(*~
	<docu>
		<summary>
			KUKA robot controller running KSS / iiQKA.OS2 9.3 (ECat).
			The interface uses 64 input and 64 output bytes. Compared to TcoKrc4 v5 it adds LocalEstopOk, NormalStop,
			CutEnableDrives, user data in both directions and a new start sequence (interface is activated first,
			drives are switched on only when CutEnableDrives is present).
		</summary>
	</docu>
~*)
FUNCTION_BLOCK TcoKukaKssEcat_v_9_3_x EXTENDS TcoIo.TcoEcatComponent IMPLEMENTS TcoAbstractions.ITcoRobotics
VAR_INPUT
    inEnable : BOOL;
END_VAR
VAR_OUTPUT
END_VAR
VAR_IN_OUT
    inoData : TcoKukaKssEcat_IO_v_9_3_x;
END_VAR
VAR
	{attribute addProperty Name "<#Status#>"}
    {attribute clr [ReadOnly()]}
    _status : TcoKukaKss_Status_v_9_3_x;
	{attribute addProperty Name "<#Control#>"}
	_control : TcoKukaKss_Control_v_9_3_x;
	{attribute addProperty Name "<#Config#>"}
    _config : TcoKukaKss_Config_v_9_3_x;
	{attribute addProperty Name "<#ECat Error#>"}
    {attribute clr [ReadOnly()]}
    _busError : BOOL;

	_someTaskIsActive : BOOL;
	_stopTasksAreActive : BOOL;

	_reportTimer : TON;
	_errorReportTimer : TON;
	{attribute 'hide'}
	_manualPV : BOOL;
END_VAR
VAR
	{attribute addProperty Name "<#Start at Main#>"}
	_startAtMainTask : TcoKukaKss_StartAtMainTask_v_9_3_x(THIS^);

	{attribute addProperty Name "<#Start motors and program#>"}
	_startMotorsAndProgramTask : TcoKukaKss_StartMotorsAndProgramTask_v_9_3_x(THIS^);

	{attribute addProperty Name "<#Start program#>"}
	_startProgramTask : TcoKukaKss_StartProgramTask_v_9_3_x(THIS^);

	{attribute addProperty Name "<#Start motors#>"}
	_startMotorsTask : TcoKukaKss_StartMotorsTask_v_9_3_x(THIS^);

	{attribute addProperty Name "<#Start movements#>"}
	_startMovementsTask : TcoKukaKss_StartMovementsTask_v_9_3_x(THIS^);

	{attribute addProperty Name "<#Start motors program and movements#>"}
	_startMotorsProgramAndMovementsTask : TcoKukaKss_StartMotorsProgramAndMovementsTask_v_9_3_x(THIS^);

	{attribute addProperty Name "<#Stop movements#>"}
	_stopMovementsTask : TcoKukaKss_StopMovementsTask_v_9_3_x(THIS^);

	{attribute addProperty Name "<#Stop movenents and program#>"}
	_stopMovementsAndProgramTask : TcoKukaKss_StopMovementsAndProgramTask_v_9_3_x(THIS^);

	{attribute addProperty Name "<#Stop program#>"}
	_stopProgramTask : TcoKukaKss_StopProgramTask_v_9_3_x(THIS^);

	{attribute addProperty Name "<#Stop motors#>"}
	_stopMotorsTask : TcoKukaKss_StopMotorsTask_v_9_3_x(THIS^);

	{attribute addProperty Name "<#Reset all outputs#>"}
	_resetAllOutputsTask : TcoKukaKss_ResetAllOutputsTask_v_9_3_x(THIS^);

    {attribute addProperty Name "<#Restore#>"}
    _restoreTask : TcoCore.TcoTask(THIS^);
END_VAR

IF NOT __ISVALIDREF(inoData) THEN
    Messenger.Post('Invalid reference', TcoCore.eMessageCategory.ProgrammingError);
    RETURN;
END_IF

SUPER^(AdsAddr := AdsAddr);
_busError := NOT SUPER^._ecatState.EcatOk;

UpdateStatus();

//MoveEnable follows the manual mode: set on entering manual mode, reset on leaving it
IF _status.State.Manual AND NOT _manualPV THEN
    _control.MoveEnable := TRUE;
ELSIF NOT _status.State.Manual AND _manualPV THEN
    _control.MoveEnable := FALSE;
END_IF
_manualPV := _status.State.Manual;

_stopTasksAreActive := _stopMovementsTask.Busy OR _stopMovementsAndProgramTask.Busy OR _stopProgramTask.Busy OR _stopMotorsTask.Busy;

_startAtMainTask.Enabled := NOT _stopTasksAreActive;
_startAtMainTask(inoConfig := _config, inoControl := _control, inoStatus := _status);

_startProgramTask.Enabled := NOT _stopTasksAreActive AND NOT _startMotorsAndProgramTask.Busy AND NOT _startMotorsTask.Busy;
_startProgramTask(inoConfig := _config, inoControl := _control, inoStatus := _status);

_startMotorsTask.Enabled := NOT _stopTasksAreActive AND NOT _startMotorsProgramAndMovementsTask.Busy AND NOT _startMotorsAndProgramTask.Busy AND NOT _startProgramTask.Busy;
_startMotorsTask(inoConfig := _config, inoControl := _control, inoStatus := _status);

_startMotorsAndProgramTask.Enabled := NOT _stopTasksAreActive AND NOT _startProgramTask.Busy AND NOT _startMotorsTask.Busy;
_startMotorsAndProgramTask(inoConfig := _config, inoControl := _control, inoStatus := _status);

_startMovementsTask.Enabled := NOT _startMotorsProgramAndMovementsTask.Busy AND NOT _stopMotorsTask.Busy;
_startMovementsTask(inoConfig := _config, inoControl := _control, inoStatus := _status);

_startMotorsProgramAndMovementsTask.Enabled := NOT _startMovementsTask.Busy AND NOT _stopMotorsTask.Busy;
_startMotorsProgramAndMovementsTask(refStartMotorsAndProgramTask := _startMotorsAndProgramTask,
    inoConfig := _config,
    inoControl := _control,
    inoStatus := _status);

_stopMovementsTask.Enabled := TRUE;
_stopMovementsTask(inoConfig := _config, inoControl := _control, inoStatus := _status);

_stopMotorsTask.Enabled := TRUE;
_stopMotorsTask(inoConfig := _config, inoControl := _control, inoStatus := _status);

_stopProgramTask.Enabled := TRUE;
_stopProgramTask(inoConfig := _config, inoControl := _control, inoStatus := _status);

_stopMovementsAndProgramTask.Enabled := TRUE;
_stopMovementsAndProgramTask(inoConfig := _config, inoControl := _control, inoStatus := _status);

_someTaskIsActive := _startAtMainTask.Busy OR
    _startProgramTask.Busy OR
    _startMotorsTask.Busy OR
    _startMotorsAndProgramTask.Busy OR
    _startMovementsTask.Busy OR
    _startMotorsProgramAndMovementsTask.Busy OR
    _stopMovementsTask.Busy OR
    _stopMovementsAndProgramTask.Busy OR
    _stopProgramTask.Busy OR
    _stopMotorsTask.Busy;

_resetAllOutputsTask.Enabled := NOT _someTaskIsActive;
_resetAllOutputsTask(inoConfig := _config, inoControl := _control, inoStatus := _status);

//*************RESTORE********************
_restoreTask.Enabled := TRUE;
IF _restoreTask.Execute() THEN
    Restore();
    _restoreTask.DoneWhen(TRUE);
END_IF
//****************************************

//do not publish diagnostic message when component is not used
IF _someTaskIsActive THEN
    IF NOT _status.State.AlarmStopActive THEN
        Messenger.Error('<#Emergency stop active#>');
    END_IF;
    IF NOT _status.State.LocalEstopOk THEN
        Messenger.Error('<#Local emergency stop active#>');
    END_IF;
    IF NOT _status.State.UserSafetySwitchClosed THEN
        Messenger.Warning('<#Safety Error #>');
    END_IF;
END_IF;

_errorReportTimer(IN := _status.State.Error, PT := _config.InfoTime);
Messenger.OnCondition(_errorReportTimer.Q).Error(_sb.Clear()
        .Append('<#Robot reported an error: #>')
        .Append(UDINT_TO_STRING(_status.State.EventId))
        .Append(' |[[0]AdvancedDiagnosticMessage]|')
        .Append('.')
        .Append('For details see the service mode')
        .ToString());

_reportTimer(IN := _status.State.Manual, PT := _config.InfoTime);
Messenger.OnCondition(_reportTimer.Q).Warning('<#Robot in manual mode. MoveEnable is set on entering manual mode!#>');

UpdateControl();

(*~
	<docu>
		<summary>
			Gets the configuration of the robot. 					
		</summary>			
	</docu>	
~*)
PROPERTY Config : REFERENCE TO TcoKukaKss_Config_v_9_3_x
GET
Config REF= _config;
END_GET
END_PROPERTY

PROPERTY PUBLIC Control : REFERENCE TO TcoKukaKss_Control_v_9_3_x
GET
Control REF= _control;
END_GET
END_PROPERTY

(*~
	<docu>
		<summary>
			Gets the status of the robot. 					
		</summary>			
	</docu>	
~*)
PROPERTY Status : REFERENCE TO TcoKukaKss_Status_v_9_3_x
GET
Status REF= _status;
END_GET
END_PROPERTY

METHOD FB_init : BOOL
VAR_INPUT
	bInitRetains : BOOL; // if TRUE, the retain variables are initialized (warm start / cold start)
	bInCopyCode : BOOL;  // if TRUE, the instance afterwards gets moved into the copy code (online change)
  	ParentObject : ITcoObject;	
END_VAR
END_METHOD

(*~
	<docu>
		<summary>
			Restores this instance to the Ready state. Can be called explicitly or from within one of the restore mechanisms.	
		</summary>			
	</docu>	
~*)
METHOD Restore : ITcoRestorable
RestoreTasks();

_control.GlobalSpeed := 0;
_control.ActivateInterface := FALSE;
_control.ErrorConfirmation := FALSE;
_control.ExternalStart := FALSE;
_control.MasterMode := 0;
_control.ToolNo := 0;
_control.WorkobjectNo := 0;
_control.PointNo := 0;
_control.UserSpecSpeed1 := 0;
_control.UserSpecSpeed2 := 0;
_control.Coordinates.X := 0;
_control.Coordinates.Y := 0;
_control.Coordinates.Z := 0;
_control.Coordinates.Rx := 0;
_control.Coordinates.Ry := 0;
_control.Coordinates.Rz := 0;
END_METHOD

METHOD INTERNAL RestoreTasks
_startAtMainTask.Restore();
_startMotorsAndProgramTask.Restore();
_startProgramTask.Restore();
_startMotorsTask.Restore();
_startMovementsTask.Restore();
_startMotorsProgramAndMovementsTask.Restore();
_stopMovementsTask.Restore();
_stopMovementsAndProgramTask.Restore();
_stopProgramTask.Restore();
_stopMotorsTask.Restore();
_resetAllOutputsTask.Restore();
END_METHOD

(*~
	<docu>
		<summary>
		    Custom service (manual, maintenance) logic.
			This method must be implemented in derived class.
		</summary>			
	</docu>	
~*)
METHOD PROTECTED ServiceMode
END_METHOD

METHOD PUBLIC StartAtMain : TcoCore.ITcoTaskStatus
StartAtMain := _startAtMainTask.Invoke();
END_METHOD

PROPERTY StartAtMainTask : TcoCore.ITcoTaskStatus
GET
StartAtMainTask := _startAtMainTask;
END_GET
END_PROPERTY

METHOD PUBLIC StartMotors : TcoCore.ITcoTaskStatus
StartMotors := _startMotorsTask.Invoke();
END_METHOD

PROPERTY StartMotorsTask : TcoCore.ITcoTaskStatus
GET
StartMotorsTask := _startMotorsTask;
END_GET
END_PROPERTY

METHOD PUBLIC StartMotorsAndProgram : TcoCore.ITcoTaskStatus
StartMotorsAndProgram := _startMotorsAndProgramTask.Invoke();
END_METHOD

PROPERTY StartMotorsAndProgramTask : TcoCore.ITcoTaskStatus
GET
StartMotorsAndProgramTask := _startMotorsAndProgramTask;
END_GET
END_PROPERTY

METHOD PUBLIC StartProgram : TcoCore.ITcoTaskStatus
StartProgram := _startProgramTask.Invoke();
END_METHOD

PROPERTY StartProgramTask : TcoCore.ITcoTaskStatus
GET
StartProgramTask := _startProgramTask;
END_GET
END_PROPERTY

METHOD PUBLIC StartMovements : TcoCore.ITcoTaskStatus
VAR_INPUT
	inData : TcoRoboticsMovementsParams;
END_VAR
StartMovements := _startMovementsTask.InvokeWithParams(inData);
END_METHOD

PROPERTY StartMovementsTask : TcoCore.ITcoTaskStatus
GET
StartMovementsTask := _startMovementsTask;
END_GET
END_PROPERTY

METHOD PUBLIC StartMotorsProgramAndMovements : TcoCore.ITcoTaskStatus
VAR_INPUT
	inData : TcoRoboticsMovementsParams;
END_VAR
StartMotorsProgramAndMovements := _startMotorsProgramAndMovementsTask.InvokeWithParams(inData);
END_METHOD

PROPERTY StartMotorsProgramAndMovementsTask : TcoCore.ITcoTaskStatus
GET
StartMotorsProgramAndMovementsTask := _startMotorsProgramAndMovementsTask;
END_GET
END_PROPERTY

METHOD PUBLIC StopMotors : TcoCore.ITcoTaskStatus
StopMotors := _stopMotorsTask.Invoke();
END_METHOD

PROPERTY StopMotorsTask : TcoCore.ITcoTaskStatus
GET
StopMotorsTask := _stopMotorsTask;
END_GET
END_PROPERTY

METHOD PUBLIC StopMovements : TcoCore.ITcoTaskStatus
VAR_INPUT
	inStopType : eTcoRoboticsStopType;
END_VAR
StopMovements := _stopMovementsTask.InvokeWithParams(inStopType);
END_METHOD

PROPERTY StopMovementsTask : TcoCore.ITcoTaskStatus
GET
StopMovementsTask := _stopMovementsTask;
END_GET
END_PROPERTY

METHOD PUBLIC StopMovementsAndProgram : TcoCore.ITcoTaskStatus
VAR_INPUT
	inStopType : eTcoRoboticsStopType;
END_VAR
StopMovementsAndProgram := _stopMovementsAndProgramTask.InvokeWithParams(inStopType);
END_METHOD

PROPERTY StopMovementsAndProgramTask : TcoCore.ITcoTaskStatus
GET
StopMovementsAndProgramTask := _stopMovementsAndProgramTask;
END_GET
END_PROPERTY

METHOD PUBLIC StopProgram : TcoCore.ITcoTaskStatus
StopProgram := _stopProgramTask.Invoke();
END_METHOD

PROPERTY StopProgramTask : TcoCore.ITcoTaskStatus
GET
StopProgramTask := _stopProgramTask;
END_GET
END_PROPERTY

METHOD PUBLIC ResetAllOutputs : TcoCore.ITcoTaskStatus
ResetAllOutputs := _resetAllOutputsTask.Invoke();
END_METHOD

PROPERTY ResetAllOutputsTask : TcoCore.ITcoTaskStatus
GET
ResetAllOutputsTask := _resetAllOutputsTask;
END_GET
END_PROPERTY

METHOD INTERNAL UpdateControl
VAR
	index : INT;
END_VAR
//SYSTEM OUTPUTS
index:=0;
inoData.Out.Outputs[index].0 := _control.ExternalStart;
inoData.Out.Outputs[index].1 := _control.MoveEnable;
inoData.Out.Outputs[index].2 := _control.ErrorConfirmation;
inoData.Out.Outputs[index].3 := _control.DrivesOff;
inoData.Out.Outputs[index].4 := _control.DrivesOn;
inoData.Out.Outputs[index].5 := _control.ActivateInterface;
inoData.Out.Outputs[index].6 := _control.StartAtMain;
inoData.Out.Outputs[index].7 := FALSE;
index:=1;
inoData.Out.Outputs[index] := 0;

//Tool signals
index:=2;
inoData.Out.Outputs[index].0 := _control.Tool_1_Retract;
inoData.Out.Outputs[index].1 := _control.Tool_1_Extend;
inoData.Out.Outputs[index].2 := _control.Tool_2_Retract;
inoData.Out.Outputs[index].3 := _control.Tool_2_Extend;
inoData.Out.Outputs[index].4 := _control.Tool_3_Retract;
inoData.Out.Outputs[index].5 := _control.Tool_3_Extend;
inoData.Out.Outputs[index].6 := _control.Tool_4_Retract;
inoData.Out.Outputs[index].7 := _control.Tool_4_Extend;
//master mode such as manual/auto ....
index:=3;
inoData.Out.Outputs[index] := _control.MasterMode;
//zone
index:=5;
inoData.Out.Outputs[index] := _control.Zone;
//position
index:=6;
inoData.Out.Outputs[index] := _control.InPosition;

//Movement parameters
index:=7;
inoData.Out.Outputs[index] := _control.ActionNo;
index:=8;
inoData.Out.Outputs[index] := _control.GlobalSpeed;
index:=9;
inoData.Out.Outputs[index] := _control.ToolNo;
index:=10;
inoData.Out.Outputs[index] := _control.WorkobjectNo;
index:=11;
inoData.Out.Outputs[index] := _control.PointNo;
index:=12;
TcoUtilities.TcoDintToBytes(inFormat:=TcoUtilities.eTcoDataFormat.LittleEndian,
							inValue:=REAL_TO_DINT(_control.UserSpecSpeed1),
							outByte0:=inoData.Out.Outputs[index],
							outByte1:=inoData.Out.Outputs[index+1],
							outByte2:=inoData.Out.Outputs[index+2],
							outByte3:=inoData.Out.Outputs[index+3]);
index:=16;
TcoUtilities.TcoDintToBytes(inFormat:=TcoUtilities.eTcoDataFormat.LittleEndian,
							inValue:=REAL_TO_DINT(_control.UserSpecSpeed2),
							outByte0:=inoData.Out.Outputs[index],
							outByte1:=inoData.Out.Outputs[index+1],
							outByte2:=inoData.Out.Outputs[index+2],
							outByte3:=inoData.Out.Outputs[index+3]);

//Coordinates
index:=20;
TcoUtilities.TcoDintToBytes(inFormat:=TcoUtilities.eTcoDataFormat.LittleEndian,
							inValue:=REAL_TO_DINT(_control.Coordinates.X * 10000.0),
							outByte0:=inoData.Out.Outputs[index],
							outByte1:=inoData.Out.Outputs[index+1],
							outByte2:=inoData.Out.Outputs[index+2],
							outByte3:=inoData.Out.Outputs[index+3]);
index:=24;
TcoUtilities.TcoDintToBytes(inFormat:=TcoUtilities.eTcoDataFormat.LittleEndian,
							inValue:=REAL_TO_DINT(_control.Coordinates.Y * 10000.0),
							outByte0:=inoData.Out.Outputs[index],
							outByte1:=inoData.Out.Outputs[index+1],
							outByte2:=inoData.Out.Outputs[index+2],
							outByte3:=inoData.Out.Outputs[index+3]);
index:=28;
TcoUtilities.TcoDintToBytes(inFormat:=TcoUtilities.eTcoDataFormat.LittleEndian,
							inValue:=REAL_TO_DINT(_control.Coordinates.Z * 10000.0),
							outByte0:=inoData.Out.Outputs[index],
							outByte1:=inoData.Out.Outputs[index+1],
							outByte2:=inoData.Out.Outputs[index+2],
							outByte3:=inoData.Out.Outputs[index+3]);
index:=32;
TcoUtilities.TcoDintToBytes(inFormat:=TcoUtilities.eTcoDataFormat.LittleEndian,
							inValue:=REAL_TO_DINT(_control.Coordinates.Rx * 10000.0),
							outByte0:=inoData.Out.Outputs[index],
							outByte1:=inoData.Out.Outputs[index+1],
							outByte2:=inoData.Out.Outputs[index+2],
							outByte3:=inoData.Out.Outputs[index+3]);
index:=36;
TcoUtilities.TcoDintToBytes(inFormat:=TcoUtilities.eTcoDataFormat.LittleEndian,
							inValue:=REAL_TO_DINT(_control.Coordinates.Ry * 10000.0),
							outByte0:=inoData.Out.Outputs[index],
							outByte1:=inoData.Out.Outputs[index+1],
							outByte2:=inoData.Out.Outputs[index+2],
							outByte3:=inoData.Out.Outputs[index+3]);
index:=40;
TcoUtilities.TcoDintToBytes(inFormat:=TcoUtilities.eTcoDataFormat.LittleEndian,
							inValue:=REAL_TO_DINT(_control.Coordinates.Rz * 10000.0),
							outByte0:=inoData.Out.Outputs[index],
							outByte1:=inoData.Out.Outputs[index+1],
							outByte2:=inoData.Out.Outputs[index+2],
							outByte3:=inoData.Out.Outputs[index+3]);

//User data from PLC to robot
FOR index := 0 TO 19 DO
	inoData.Out.Outputs[44 + index] := _control.DataToRobot[index];
END_FOR
END_METHOD

METHOD INTERNAL UpdateStatus
VAR
	index : INT;
	_bytes : DINT;
END_VAR
//SYSTEM INPUTS
index:=0;
_status.State.RcReady := inoData.In.Inputs[index].0;
_status.State.AlarmStopActive := inoData.In.Inputs[index].1;
_status.State.UserSafetySwitchClosed := inoData.In.Inputs[index].2;
_status.State.DrivesReady := inoData.In.Inputs[index].3;
_status.State.RobotCalibrated := inoData.In.Inputs[index].4;
_status.State.InterfaceActivated := inoData.In.Inputs[index].5;
_status.State.StopMess := inoData.In.Inputs[index].6;
_status.State.RobotStopped := inoData.In.Inputs[index].7;

index:=1;
_status.State.InHome := inoData.In.Inputs[index].0;
_status.State.Manual := inoData.In.Inputs[index].1;
_status.State.LocalEstopOk := inoData.In.Inputs[index].2;
_status.State.ExternalAutomatic := inoData.In.Inputs[index].3;
_status.State.ProActive := inoData.In.Inputs[index].4;
_status.State.PpMoved := inoData.In.Inputs[index].5;
_status.State.Error := inoData.In.Inputs[index].6;
_status.State.ProgramMoveActive := inoData.In.Inputs[index].7;

//Area/positions flags this should be obsolete because Zones and InPosition is used as byte below
index:=2;
_status.State.InArea_1 := inoData.In.Inputs[index].0;
_status.State.InArea_2 := inoData.In.Inputs[index].1;
_status.State.InArea_3 := inoData.In.Inputs[index].2;
_status.State.InArea_4 := inoData.In.Inputs[index].3;
_status.State.InPosition_1 := inoData.In.Inputs[index].4;
_status.State.InPosition_2 := inoData.In.Inputs[index].5;
_status.State.InPosition_3 := inoData.In.Inputs[index].6;
_status.State.InPosition_4 := inoData.In.Inputs[index].7;

//Tool signals
index:=3;
_status.State.Tool_1_Retract := inoData.In.Inputs[index].0;
_status.State.Tool_1_Extend := inoData.In.Inputs[index].1;
_status.State.Tool_2_Retract := inoData.In.Inputs[index].2;
_status.State.Tool_2_Extend := inoData.In.Inputs[index].3;
_status.State.Tool_3_Retract := inoData.In.Inputs[index].4;
_status.State.Tool_3_Extend := inoData.In.Inputs[index].5;
_status.State.Tool_4_Retract := inoData.In.Inputs[index].6;
_status.State.Tool_4_Extend := inoData.In.Inputs[index].7;

//Normal stop / drives enable (KSS 9.3)
index:=4;
_status.State.NormalStop := inoData.In.Inputs[index].0;
_status.State.CutEnableDrives := inoData.In.Inputs[index].1;

index:=5;
_status.State.Zone := inoData.In.Inputs[index];
index:=6;
_status.State.InPosition := inoData.In.Inputs[index];

//Movement parameters
index:=7;
_status.State.ActionNo := inoData.In.Inputs[index];
index:=8;
_status.State.GlobalSpeed := inoData.In.Inputs[index];
index:=9;
_status.State.ToolNo := inoData.In.Inputs[index];
index:=10;
_status.State.WorkobjectNo := inoData.In.Inputs[index];
index:=11;
_status.State.PointNo := inoData.In.Inputs[index];
index:=12;
_status.State.UserSpecSpeed1 := TcoUtilities.TcoBytesToDint(inFormat:=TcoUtilities.eTcoDataFormat.LittleEndian,
							inByte0:=inoData.In.Inputs[index],
							inByte1:=inoData.In.Inputs[index+1],
							inByte2:=inoData.In.Inputs[index+2],
							inByte3:=inoData.In.Inputs[index+3]);
index:=16;
_status.State.UserSpecSpeed2 := TcoUtilities.TcoBytesToDint(inFormat:=TcoUtilities.eTcoDataFormat.LittleEndian,
							inByte0:=inoData.In.Inputs[index],
							inByte1:=inoData.In.Inputs[index+1],
							inByte2:=inoData.In.Inputs[index+2],
							inByte3:=inoData.In.Inputs[index+3]);
index:=20;
_bytes := TcoUtilities.TcoBytesToDint(inFormat:=TcoUtilities.eTcoDataFormat.LittleEndian,
							inByte0:=inoData.In.Inputs[index],
							inByte1:=inoData.In.Inputs[index+1],
							inByte2:=inoData.In.Inputs[index+2],
							inByte3:=inoData.In.Inputs[index+3]);
_status.State.Coordinates.X := DINT_TO_REAL(_bytes) / 10000.0;

index:=24;
_bytes := TcoUtilities.TcoBytesToDint(inFormat:=TcoUtilities.eTcoDataFormat.LittleEndian,
							inByte0:=inoData.In.Inputs[index],
							inByte1:=inoData.In.Inputs[index+1],
							inByte2:=inoData.In.Inputs[index+2],
							inByte3:=inoData.In.Inputs[index+3]);
_status.State.Coordinates.Y := DINT_TO_REAL(_bytes) / 10000.0;

index:=28;
_bytes := TcoUtilities.TcoBytesToDint(inFormat:=TcoUtilities.eTcoDataFormat.LittleEndian,
							inByte0:=inoData.In.Inputs[index],
							inByte1:=inoData.In.Inputs[index+1],
							inByte2:=inoData.In.Inputs[index+2],
							inByte3:=inoData.In.Inputs[index+3]);
_status.State.Coordinates.Z := DINT_TO_REAL(_bytes) / 10000.0;

index:=32;
_bytes := TcoUtilities.TcoBytesToDint(inFormat:=TcoUtilities.eTcoDataFormat.LittleEndian,
							inByte0:=inoData.In.Inputs[index],
							inByte1:=inoData.In.Inputs[index+1],
							inByte2:=inoData.In.Inputs[index+2],
							inByte3:=inoData.In.Inputs[index+3]);
_status.State.Coordinates.Rx := DINT_TO_REAL(_bytes) / 10000.0;

index:=36;
_bytes := TcoUtilities.TcoBytesToDint(inFormat:=TcoUtilities.eTcoDataFormat.LittleEndian,
							inByte0:=inoData.In.Inputs[index],
							inByte1:=inoData.In.Inputs[index+1],
							inByte2:=inoData.In.Inputs[index+2],
							inByte3:=inoData.In.Inputs[index+3]);
_status.State.Coordinates.Ry := DINT_TO_REAL(_bytes) / 10000.0;

index:=40;
_bytes := TcoUtilities.TcoBytesToDint(inFormat:=TcoUtilities.eTcoDataFormat.LittleEndian,
							inByte0:=inoData.In.Inputs[index],
							inByte1:=inoData.In.Inputs[index+1],
							inByte2:=inoData.In.Inputs[index+2],
							inByte3:=inoData.In.Inputs[index+3]);
_status.State.Coordinates.Rz := DINT_TO_REAL(_bytes) / 10000.0;

index:=44;
_status.State.EventId := TcoUtilities.TcoBytesToUDint(inFormat:=TcoUtilities.eTcoDataFormat.LittleEndian,
							inByte0:=inoData.In.Inputs[index],
							inByte1:=inoData.In.Inputs[index+1],
							inByte2:=inoData.In.Inputs[index+2],
							inByte3:=inoData.In.Inputs[index+3]);

//User data from robot to PLC
FOR index := 0 TO 15 DO
	_status.State.DataFromRobot[index] := inoData.In.Inputs[48 + index];
END_FOR
END_METHOD

END_FUNCTION_BLOCK

(* stored: Version 1.1.0.1, ProductVersion 3.1.4024.12
   POU TcoKukaKssEcat_v_9_3_x: Id {8240f261-28f6-44a7-bcaa-32d5ed3116a8}, SpecialFunc None
   Folder Operations: Id {027f61ae-e71f-4a4c-8c22-228286bc5d5f}
   Folder Task: Id {2c37f829-6297-4777-bc3f-0fc886118850}
   Property Config: Id {4d37f924-eb41-4fef-9edc-76d0b4f40692}
   Get Get: Id {2258dc20-4fdb-45fe-b63a-6505710d1a93}
   Property Control: Id {e3180703-86e2-43b3-b541-81614d7caa3a}
   Get Get: Id {5ec5fc1e-f975-4259-ba8d-465a1bce42c6}
   Property Status: Id {aecf7611-2d37-4ec3-914d-10b4282d2e15}
   Get Get: Id {f0ec804c-6393-401c-a4aa-7a6926518852}
   Method FB_init: Id {84391af5-c8c2-48d5-aef9-953e5348a8cc}
   Method Restore: Id {a1cbd8ee-e5e1-46f7-af77-87e7a40f6df0}
   Method RestoreTasks: Id {9d5410f7-dc53-40b8-a734-97bf164b14c6}
   Method ServiceMode: Id {70f72e03-0c48-49f2-978d-d8c5f04bad64}
   Method StartAtMain: Id {ee26d6c3-6987-4325-9ae8-9935b48b6916}
   Property StartAtMainTask: Id {0e9a2e65-9ea4-424f-8aaa-4bbac75b198b}
   Get Get: Id {1daf6033-70d9-4fa3-958c-664cd6aec491}
   Method StartMotors: Id {80517a4e-2da5-4a09-9eb2-dcf97517ae03}
   Property StartMotorsTask: Id {f0764713-c55f-4e98-92c4-76446bc58f88}
   Get Get: Id {e58a6284-6ff5-43cb-ba0e-5bdf3165ede0}
   Method StartMotorsAndProgram: Id {92cb27c3-6fe5-4c79-b4db-a5fcb2c6cc1b}
   Property StartMotorsAndProgramTask: Id {6f675b0f-81cf-4ece-82b8-033f789339dd}
   Get Get: Id {8bbeb0b0-08e6-4080-b0b1-c84f245e676e}
   Method StartProgram: Id {ae2183a9-10ad-403e-981c-3accd56196b6}
   Property StartProgramTask: Id {5e8f02c7-d1e2-4f65-8121-1ca5dfda42f3}
   Get Get: Id {95d71a20-792e-4399-b0b3-def447abee8f}
   Method StartMovements: Id {e0e903ef-2eca-4f60-bcbb-8b7c8eb2a44b}
   Property StartMovementsTask: Id {a253a85d-c4be-4ced-82a8-ed8b22f987a4}
   Get Get: Id {d3400dcb-fbca-4a9f-9c49-3655ace27497}
   Method StartMotorsProgramAndMovements: Id {9f9204f3-ee20-43f0-9e7f-cee360d91101}
   Property StartMotorsProgramAndMovementsTask: Id {f6e52590-e9ee-4e95-852f-ff595d460baf}
   Get Get: Id {0fd75fcf-1e92-44c1-99a4-d9e5737ab122}
   Method StopMotors: Id {d39b24d0-0671-483d-a65a-e48964909436}
   Property StopMotorsTask: Id {1ad48295-fd68-4185-9029-35145454f32e}
   Get Get: Id {902949f0-48ca-4d6e-b91c-1a7a13dda50f}
   Method StopMovements: Id {ce5e2a94-a8ff-45ae-948e-3fec922d2198}
   Property StopMovementsTask: Id {907c6652-6f82-4a9d-9fc2-d5bb2e6a1457}
   Get Get: Id {dd059e4e-b76a-4df0-81db-453fe42ccb9a}
   Method StopMovementsAndProgram: Id {0d63daf9-9853-46f7-9c05-f2e8fa40f56d}
   Property StopMovementsAndProgramTask: Id {98da0b98-1a57-4831-bc2c-cc80cb53abdc}
   Get Get: Id {baa163a4-d513-4e44-bd7a-8eb973a5c095}
   Method StopProgram: Id {a09c42a3-d31b-4a6e-acc8-82b54db96d96}
   Property StopProgramTask: Id {fb272975-8f2d-45c3-9fa3-0005671b3436}
   Get Get: Id {8f4df811-2057-426e-aecb-8e1a5c6f93c8}
   Method ResetAllOutputs: Id {8b395219-0402-441e-ba4f-854d2840fd1b}
   Property ResetAllOutputsTask: Id {516753eb-66dd-4c02-80eb-73b687ead365}
   Get Get: Id {47a28248-e34b-4eca-9921-12cbb19cc271}
   Method UpdateControl: Id {278e97c0-beba-48d8-87f8-eb708cd7d52c}
   Method UpdateStatus: Id {9e075e75-089b-4b26-b7b0-8a85eb16f24c} *)
